// Mitsubishi GX Works2 project: 261012_타이머실습_일반타이머고속   PLC: Q03UDV

PROGRAM MAIN
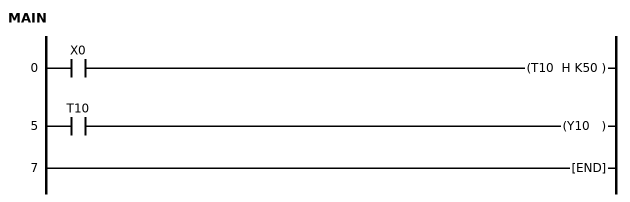
0     LD      X0
      OUTH    T10 K50
5     LD      T10
      OUT     Y10
7     END
END_PROGRAM
